Fanuc KAREL source: KA00082.KL

PROGRAM KA00082
%NOLOCKGROUP
VAR
  SRC: XYZWPREXT
  DST: CONFIG
BEGIN
  SRC.X = 1.0
  DST = SRC
END KA00082
